(* IEC 61131-3 sources: s7-to-codesys/tests/POUs/S7Compat/FB_S7Ton_Test, 8 files *)

(* ---- FB_S7Ton_Test.decl.st ---- *)
// Назначение: набор тестов CfUnit (coUnit 1.2.0.0) для FB_S7Ton слоя совместимости S7Compat:
//             отсчёт с фронта IN и с первого вызова при IN = TRUE, Q ровно на пороге PT, насыщение
//             ET, сброс по IN = FALSE, PT = 0, переход TIME через 2^32 мс (в том числе Q при IN = TRUE
//             дольше 2^32 мс), совпадение со Standard.TON в реальном времени (тест на несколько циклов).
//             Ожидаемые значения — по семантике МЭК 61131-3 и S7 (описание в объявлении блока), а
//             не по результату реализации. Моделируемое время — GVL_S7Clock (тест включает и
//             выключает его сам). Экземпляр набора объявляется в PRG_Tests.
// Автор:      kr0nsch
// Версия:     0.1.0
// Документ:   docs/methodology.md, раздел «Проверка поведения: время в тестах»
FUNCTION_BLOCK FB_S7Ton_Test EXTENDS coUnit.FB_TestSuite
VAR
    // MatchesStandardInRealTime: состояние между циклами (тест идёт несколько циклов)
    fbRtCompat : FB_S7Ton;              // проверяемый таймер S7Compat
    fbRtStandard : TON;               // эталон — таймер CODESYS Standard
    xRtStarted : BOOL;              // момент начала зафиксирован
    xRtDone : BOOL;                 // тест завершён
    xRtIn : BOOL;                   // общий вход IN
    xRtSawQ : BOOL;                 // Standard Q хотя бы раз был TRUE
    tRtStart : TIME;                // время начала теста (F_S7Now() = TIME())
    tRtElapsed : TIME;              // прошло с начала теста
    tRtEtDiff : TIME;               // |ET S7Compat - ET Standard|
    tRtEtToPt : TIME;               // PT - ET Standard (близость к порогу)
    iRtMismatches : INT;            // циклов с расхождением
END_VAR
VAR CONSTANT
    T_RT_PT : TIME := T#200MS;      // PT обоих таймеров
    T_RT_DURATION : TIME := T#700MS;  // длительность теста
    T_RT_TOL : TIME := T#5MS;       // допуск ET: таймеры читают TIME() в разные моменты цикла
END_VAR

(* ---- CountsFromRisingEdge.method.decl.st ---- *)
// IN = TRUE с t = 1000 мс, PT = 2 с: Q = FALSE до 2999 мс, TRUE ровно на 3000 мс; ET растёт до PT и стоит.
METHOD PRIVATE CountsFromRisingEdge
VAR
    fbDut : FB_S7Ton;       // проверяемый таймер (новый экземпляр на каждый вызов метода)
END_VAR

(* ---- FirstCallWithInTrueStarts.method.decl.st ---- *)
// первый вызов экземпляра уже с IN = TRUE (t = 500 мс) — начало отсчёта.
METHOD PRIVATE FirstCallWithInTrueStarts
VAR
    fbDut : FB_S7Ton;       // проверяемый таймер (новый экземпляр на каждый вызов метода)
END_VAR

(* ---- KeepsQWhileInHeldAcrossWrap.method.decl.st ---- *)
// IN = TRUE без перерыва дольше 2^32 мс (около 49,7 суток): Q не падает после перехода TIME через ноль — в S7
// и у Standard.TON Q держится, пока IN = TRUE. Разность «сейчас − старт» по модулю 2^32 здесь неверна:
// прошло 2^32 + 396 мс, а разность — 100 мс.
METHOD PRIVATE KeepsQWhileInHeldAcrossWrap
VAR
    fbDut : FB_S7Ton;       // проверяемый таймер (новый экземпляр на каждый вызов метода)
END_VAR

(* ---- MatchesStandardInRealTime.method.impl.st ---- *)
coUnit.TEST('MatchesStandardInRealTime');
IF NOT xRtDone THEN
    IF NOT xRtStarted THEN
        xRtStarted := TRUE;
        tRtStart := F_S7Now();  // xSimulation = FALSE: время ПЛК, как TIME()
    END_IF
    tRtElapsed := F_S7Now() - tRtStart;
    xRtIn := (tRtElapsed < T#300MS) OR (tRtElapsed >= T#400MS AND tRtElapsed < T#520MS);
    fbRtCompat(IN := xRtIn, PT := T_RT_PT);
    fbRtStandard(IN := xRtIn, PT := T_RT_PT);
    IF fbRtCompat.ET >= fbRtStandard.ET THEN
        tRtEtDiff := fbRtCompat.ET - fbRtStandard.ET;
    ELSE
        tRtEtDiff := fbRtStandard.ET - fbRtCompat.ET;
    END_IF
    tRtEtToPt := T_RT_PT - fbRtStandard.ET;  // ET <= PT
    IF tRtEtDiff > T_RT_TOL OR (fbRtCompat.Q <> fbRtStandard.Q AND tRtEtToPt > T_RT_TOL) THEN
        iRtMismatches := iRtMismatches + 1;
    END_IF
    xRtSawQ := xRtSawQ OR fbRtStandard.Q;
    IF tRtElapsed >= T_RT_DURATION THEN
        xRtDone := TRUE;
        AssertEquals_INT(Expected := 0, Actual := iRtMismatches, Message := 'FB_S7Ton vs TON: mismatching cycles');
        AssertTrue(Condition := xRtSawQ, Message := 'FB_S7Ton vs TON: Standard Q never TRUE, test did not run');
    END_IF
END_IF
IF xRtDone THEN
    coUnit.TEST_FINISHED();
END_IF

(* ---- ResetWhenInFalse.method.decl.st ---- *)
// IN = FALSE сбрасывает Q и ET; новый фронт — отсчёт заново.
METHOD PRIVATE ResetWhenInFalse
VAR
    fbDut : FB_S7Ton;       // проверяемый таймер (новый экземпляр на каждый вызов метода)
END_VAR

(* ---- SurvivesTimeWraparound.method.decl.st ---- *)
// переход TIME через 2^32 мс (около 49,7 суток): разность моментов — по модулю 2^32.
METHOD PRIVATE SurvivesTimeWraparound
VAR
    fbDut : FB_S7Ton;       // проверяемый таймер (новый экземпляр на каждый вызов метода)
END_VAR

(* ---- ZeroPtSwitchesImmediately.method.decl.st ---- *)
// PT = 0: Q = TRUE уже на вызове с фронтом IN (прошло 0 >= 0).
METHOD PRIVATE ZeroPtSwitchesImmediately
VAR
    fbDut : FB_S7Ton;       // проверяемый таймер (новый экземпляр на каждый вызов метода)
END_VAR
